{attribute 'qualified_only'}
{attribute 'strict'}
{attribute 'to_string'}
TYPE E_USint :
(
	eOptionA := 0,
	eOptionB,
	eOptionC
) USINT;
END_TYPE

(* stored: Version 1.1.0.1, ProductVersion 3.1.4026.19
   DUT E_USint: Id {8b2be9b2-4670-48b4-bc0e-ffa857726f4a} *)
